(* IEC 61131-3 sources: JingjiangMoonbox/Application/Application/任务列表/公用函数, 4 files *)

(* ---- KS_GetBitByDword.st ---- *)
(*@CES
Name=KS_GetBitByDword
Type=FunctionBlock
TypeGuid=6f9dac99-8de1-4efc-8465-68ac443b7d08
Guid=6ef6fac5-03f1-4f35-a007-cccb879e1ed9
HasDeclaration=True
HasImplementation=True
*)
{DECLARATION}
FUNCTION KS_GetBitByDword : BOOL(*获取Dword中的位*)
VAR_INPUT
	i_byBitId:BYTE;(*0--31*)
	i_dwValue:DWORD;
END_VAR
VAR
	xGetDne: BOOL;
	dwTmp: DWORD;
	xBit:BOOL;
END_VAR
{IMPLEMENTATION}
IF i_byBitId>=0 AND
	i_byBitId<16 THEN
	dwTmp:=SHR(i_dwValue,i_byBitId);
	xBit:=dwTmp.0;
END_IF
KS_GetBitByDword:=xBit;

(* ---- KS_GetBitByWord.st ---- *)
(*@CES
Name=KS_GetBitByWord
Type=FunctionBlock
TypeGuid=6f9dac99-8de1-4efc-8465-68ac443b7d08
Guid=14ad4b69-ea73-4214-a3fe-9debcfa02eec
HasDeclaration=True
HasImplementation=True
*)
{DECLARATION}
FUNCTION KS_GetBitByWord : BOOL(*获取word中的位*)
VAR_INPUT
	i_byBitId:BYTE;(*0--15*)
	i_wValue:WORD;
END_VAR
VAR
	xGetDne: BOOL;
	wTmp: WORD;
	xBit:BOOL;
END_VAR
{IMPLEMENTATION}
IF i_byBitId>=0 AND
	i_byBitId<16 THEN
	wTmp:=SHR(i_wValue,i_byBitId);
	xBit:=wTmp.0;
END_IF
KS_GetBitByWord:=xBit;

(* ---- KS_MOD_LREAL.st ---- *)
(*@CES
Name=KS_MOD_LREAL
Type=FunctionBlock
TypeGuid=6f9dac99-8de1-4efc-8465-68ac443b7d08
Guid=c7df3acb-0909-4f65-9b34-010cacb37200
HasDeclaration=True
HasImplementation=True
*)
{DECLARATION}
FUNCTION KS_MOD_LREAL : LREAL(*浮点数的取模*)
VAR_INPUT
	i_lrData:LREAL;
	i_rMOD:REAL;
END_VAR
VAR
	iTimes: INT;
	iN: INT;
	lrTemp: LREAL;
END_VAR
{IMPLEMENTATION}
IF i_rMOD<>0 THEN
	iTimes:=LREAL_TO_INT(i_lrData/i_rMOD);
END_IF

lrTemp:=i_lrData-i_rMOD*iTimes;
IF lrTemp<0 THEN
	lrTemp:=lrTemp+i_rMOD;
END_IF
KS_MOD_LREAL:=lrTemp;

(* ---- KS_SetWordBit.st ---- *)
(*@CES
Name=KS_SetWordBit
Type=FunctionBlock
TypeGuid=6f9dac99-8de1-4efc-8465-68ac443b7d08
Guid=02828fa7-5c3c-4227-9d4b-97efc9023b71
HasDeclaration=True
HasImplementation=True
*)
{DECLARATION}
FUNCTION KS_SetWordBit : BOOL(*设置word位*)
VAR_INPUT
	i_byBitId:BYTE;(*0--15*)
	i_xSetBool:BOOL;
	i_pwValue:POINTER TO WORD;
END_VAR
VAR
	wTmp: WORD;
	xSetDne: BOOL;
END_VAR
{IMPLEMENTATION}
IF i_byBitId>=0 AND
	i_byBitId<16 THEN

	wTmp:=16#00000001;
	wTmp:=SHL(wTmp,i_byBitId);

	IF i_pwValue<>0 THEN
		IF i_xSetBool THEN(*写1*)
			i_pwValue^:=i_pwValue^ OR wTmp;
		ELSE(*写0*)
			wTmp:=NOT wTmp;(*先取反*)
			i_pwValue^:=i_pwValue^ AND wTmp;
		END_IF

		xSetDne:=TRUE;
	END_IF
ELSE;
END_IF
KS_SetWordBit:=xSetDne;
